(* IEC 61131-3 sources: codesys-framework/txt/application/ToDo/Hyperion/Enum, 5 files *)

(* ---- E_HyperionForceLoggingHandShake.dut.st ---- *)
TYPE E_HyperionForceLoggingHandShake :
(
	None						:= 0,
	AwaitingForceForceLogging 		:= 14,
	AwaitingClearForceLogging 		:= 15,
	AwaitingFinishForceLogging     := 16

);
END_TYPE

(* ---- E_HyperionHandshake.dut.st ---- *)
TYPE E_HyperionHandshake :
(
	Invalid := 0,
	AwaitingSendStartRqst := 1,
	AwaitingSendStopRqst := 2,
	AwaitingStartAckNack := 3,
	AwaitingStopAckNack := 4,

	Rcve_StartRqst := 5,

	Send_ReadyForStart := 6,
	Send_NotReadyForStart := 7,

	Rcve_StopRqst := 8,

	DataValidating := 9,
	Send_DataValid := 10,
	Send_DataNotValid := 11
);
END_TYPE

(* ---- E_HyperionOutputResendHandShake.dut.st ---- *)
TYPE E_HyperionOutputResendHandShake :
(
	None						:= 0,
	AwaitingForceResendOutputParam 		:= 14,
	AwaitingClearResendOutputParam 		:= 15,
	AwaitingFinishResendOutputParam     := 16

);
END_TYPE

(* ---- E_ParameterMode.dut.st ---- *)
TYPE E_ParameterMode :
(
	Invalid := 0,
	CheckHyp := 1,
	CheckPLC := 2,
	ValidateHyp := 3,
	SavePLC := 4,
	ValidateHypAndSavePLC := 5,
	CopyPLCToHyp := 6
);
END_TYPE

(* ---- E_ParameterValidationCode.dut.st ---- *)
TYPE E_ParameterValidationCode :
(
	Invalid := 0,
	Validation_Failed_IsZero := 1,
	Validation_Failed_BelowMinimum := 2,
	Validation_Failed_AboveMaximum := 3,
	Validation_Failed_External := 4,
	Validation_Ok := 5
);
END_TYPE
